(* IEC 61131-3 sources: ADRC_WWTP/PLC_ST/Codigos, 7 files *)

(* ---- ADRC_ESO.st ---- *)
FUNCTION_BLOCK ADRC_ESO
VAR_INPUT
    SET_POINT : LREAL;              (* setpoint r *)
    ACTUAL    : LREAL;              (* measurement y *)
    WC        : LREAL;              (* controller bandwidth [rad/s] *)
    WO        : LREAL;              (* observer bandwidth [rad/s] *)
    B0        : LREAL;              (* plant input gain *)
    TS        : TIME := T#50MS;     (* sampling time, equal to the task period *)
    U_MIN     : LREAL := 0.0;
    U_MAX     : LREAL := 100.0;
    RESET     : BOOL := FALSE;
END_VAR
VAR_OUTPUT
    U         : LREAL;              (* control signal to the actuator *)
END_VAR
VAR CONSTANT
    ST_RESET     : INT := 0;
    ST_AUTOMATIC : INT := 1;
END_VAR
VAR
    T_S       : LREAL;              (* sampling time [s] *)
    State     : INT;
    Ready     : BOOL := FALSE;      (* valid gains available *)
    A         : ARRAY[1..2, 1..2] OF LREAL;
    B         : ARRAY[1..2] OF LREAL;
    C         : ARRAY[1..2] OF LREAL;
    L         : ARRAY[1..2] OF LREAL;
    K         : ARRAY[1..2] OF LREAL;
    X         : ARRAY[1..2] OF LREAL;   (* x_hat: estimated error and total disturbance *)
    X_old     : ARRAY[1..2] OF LREAL;
    Ey, Ey_old : LREAL;
    U0, U0_old : LREAL;
    Bo, Zc, Zo : LREAL;
END_VAR

(* state selection *)
IF RESET OR NOT Ready THEN
    State := ST_RESET;
ELSE
    State := ST_AUTOMATIC;
END_IF

(* sampling time in seconds *)
T_S := TIME_TO_LREAL(TS) / 1000.0;

(* gains are only updated outside AUTOMATIC *)
IF (State <> ST_AUTOMATIC) AND (T_S > 0.0) AND (WC > 0.0) AND (WO > WC) AND (B0 > 0.0) THEN
    Zc := EXP(-WC * T_S);
    Zo := EXP(-WO * T_S);
    A[1,1] := 1.0;   A[1,2] := T_S;
    A[2,1] := 0.0;   A[2,2] := 1.0;
    B[1]   := T_S;    B[2]   := 0.0;
    C[1]   := 1.0;   C[2]   := 0.0;
    L[1]   := 2.0 * (1.0 - Zo);
    L[2]   := (1.0 - Zo) * (1.0 - Zo) / T_S;
    K[1]   := (1.0 - Zc) / T_S;
    K[2]   := 1.0;
    Bo     := B0;
    Ready  := TRUE;
END_IF

(* observer: x_hat[k] = (A - L C) x_hat[k-1] + B u0[k-1] + L ey[k-1] *)
X[1] := (A[1,1] - L[1]*C[1])*X_old[1] + (A[1,2] - L[1]*C[2])*X_old[2] + B[1]*U0_old + L[1]*Ey_old;
X[2] := (A[2,1] - L[2]*C[1])*X_old[1] + (A[2,2] - L[2]*C[2])*X_old[2] + B[2]*U0_old + L[2]*Ey_old;

CASE State OF
ST_RESET:
    (* output and observer to zero, as if it had just started *)
    U    := LIMIT(U_MIN, 0.0, U_MAX);
    X[1] := 0.0;
    X[2] := -Bo * U;
    Ey   := 0.0;

ST_AUTOMATIC:
    (* control law: u0 = -K x_hat[k],  u = u0/b0 *)
    Ey := ACTUAL - SET_POINT;
    U0 := -(K[1]*X[1] + K[2]*X[2]);
    U  := LIMIT(U_MIN, U0 / Bo, U_MAX);
END_CASE

(* the observer always receives the applied order *)
U0 := Bo * U;

X_old  := X;
U0_old := U0;
Ey_old := Ey;
END_FUNCTION_BLOCK

(* ---- ADRC_GPI.st ---- *)
FUNCTION_BLOCK ADRC_GPI
VAR_INPUT
    SET_POINT : LREAL;              (* setpoint r *)
    ACTUAL    : LREAL;              (* measurement y *)
    WC        : LREAL;              (* controller bandwidth [rad/s] *)
    WO        : LREAL;              (* observer bandwidth [rad/s] *)
    B0        : LREAL;              (* plant input gain *)
    TS        : TIME := T#50MS;     (* sampling time, equal to the task period *)
    U_MIN     : LREAL := 0.0;
    U_MAX     : LREAL := 100.0;
    RESET     : BOOL := FALSE;
END_VAR
VAR_OUTPUT
    U         : LREAL;              (* control signal to the actuator *)
END_VAR
VAR CONSTANT
    ST_RESET     : INT := 0;
    ST_AUTOMATIC : INT := 1;
END_VAR
VAR
    T_S       : LREAL;              (* sampling time [s] *)
    State     : INT;
    Ready     : BOOL := FALSE;      (* valid gains available *)
    Bo, D0, Q : LREAL;
    A1, A2    : LREAL;              (* common denominator of H1 and H2 *)
    B0z, B1z, B2z : LREAL;          (* numerator of H1 *)
    G0, G1, G2    : LREAL;          (* numerator of H2 *)
    E, E_1, E_2   : LREAL;          (* r - y and its delays *)
    V, V_1, V_2   : LREAL;
    U_1, U_2, W   : LREAL;
END_VAR

(* state selection *)
IF RESET OR NOT Ready THEN
    State := ST_RESET;
ELSE
    State := ST_AUTOMATIC;
END_IF

(* sampling time in seconds *)
T_S := TIME_TO_LREAL(TS) / 1000.0;

(* gains are only updated outside AUTOMATIC *)
IF (State <> ST_AUTOMATIC) AND (T_S > 0.0) AND (WC > 0.0) AND (WO > WC) AND (B0 > 0.0) THEN
    (* Tustin with E1(s) = (s + wo)^2 *)
    Q   := 2.0 + WO * T_S;
    D0  := Q * Q;
    A1  := -2.0 * (4.0 - WO * WO * T_S * T_S) / D0;
    A2  := (2.0 - WO * T_S) * (2.0 - WO * T_S) / D0;
    B0z := WO * T_S * (WC * WO * T_S + 2.0 * (WO + 2.0 * WC)) / D0;
    B1z := 2.0 * WC * WO * WO * T_S * T_S / D0;
    B2z := WO * T_S * (WC * WO * T_S - 2.0 * (WO + 2.0 * WC)) / D0;
    G0  := T_S * (2.0 * WC - WO * WO * T_S) / D0;
    G1  := -2.0 * WO * WO * T_S * T_S / D0;
    G2  := -T_S * (2.0 * WC + WO * WO * T_S) / D0;
    Bo  := B0;
    Ready := TRUE;
END_IF

CASE State OF
ST_RESET:
    (* output and delays to zero, as if it had just started *)
    U := LIMIT(U_MIN, 0.0, U_MAX);
    E := 0.0;   E_1 := 0.0;   E_2 := 0.0;
    V := U;     V_1 := U;     V_2 := U;
    U_1 := U;   U_2 := U;

ST_AUTOMATIC:
    (* direct form I; 1 + G0 solves the loop through the direct term of H2 *)
    E := SET_POINT - ACTUAL;
    W := (B0z*E + B1z*E_1 + B2z*E_2) / Bo - (G1*U_1 + G2*U_2) - A1*V_1 - A2*V_2;
    U := LIMIT(U_MIN, W / (1.0 + G0), U_MAX);
    V := W - G0 * U;
END_CASE

(* shift: oldest first *)
E_2 := E_1;   E_1 := E;
V_2 := V_1;   V_1 := V;
U_2 := U_1;   U_1 := U;
END_FUNCTION_BLOCK

(* ---- BEZIER_REF.st ---- *)
FUNCTION_BLOCK BEZIER_REF
VAR_INPUT
    SET_POINT : LREAL;              (* setpoint r *)
    ACTUAL    : LREAL;              (* measurement y *)
    TF        : TIME := T#20M;      (* segment duration, taken at each setpoint change *)
    TS        : TIME := T#50MS;     (* sampling time, equal to the task period *)
    RESET     : BOOL := FALSE;
END_VAR
VAR_OUTPUT
    Y         : LREAL;              (* reference y*, goes to the controller *)
END_VAR
VAR CONSTANT
    ST_RESET     : INT := 0;
    ST_AUTOMATIC : INT := 1;
END_VAR
VAR
    T_S       : LREAL;              (* sampling time [s] *)
    T_F       : LREAL;              (* segment duration [s] *)
    State     : INT;
    Ready     : BOOL := FALSE;      (* valid parameters available *)
    Ts_set         : LREAL;
    Tf_set         : LREAL;         (* duration of the current segment *)
    Yc, Dyc, Yf    : LREAL;         (* segment start state and target *)
    Delta, C1, C2, C3 : LREAL;      (* polynomial coefficients in tau *)
    Dy, Tn, Cnt, SP_old : LREAL;
END_VAR

(* state selection *)
IF RESET OR NOT Ready THEN
    State := ST_RESET;
ELSE
    State := ST_AUTOMATIC;
END_IF

(* times in seconds *)
T_S := TIME_TO_LREAL(TS) / 1000.0;
T_F := TIME_TO_LREAL(TF) / 1000.0;

(* parameters are only updated outside AUTOMATIC *)
IF (State <> ST_AUTOMATIC) AND (T_S > 0.0) AND (T_F > 0.0) THEN
    Ts_set := T_S;
    Tf_set := T_F;
    Ready  := TRUE;
END_IF

CASE State OF
ST_RESET:
    (* at rest on the measurement; leaving RESET starts the manoeuvre again *)
    Y  := ACTUAL;   Dy := 0.0;
    Yc := ACTUAL;   Dyc := 0.0;   Yf := ACTUAL;
    C1 := 0.0;      C2 := 0.0;    C3 := 0.0;
    Cnt := 0.0;     SP_old := ACTUAL;

ST_AUTOMATIC:
    (* evaluate the current segment, tau = n Ts/Tf *)
    Tn := Cnt * Ts_set / Tf_set;
    IF Tn < 1.0 THEN
        Y  := Yc + Tn * (C1 + Tn * (C2 + Tn * C3));
        Dy := (C1 + Tn * (2.0 * C2 + 3.0 * Tn * C3)) / Tf_set;
    ELSE
        Y  := Yf;
        Dy := 0.0;
    END_IF

    (* new setpoint: replan from the state of the reference *)
    IF SET_POINT <> SP_old THEN
        Yc := Y;
        Dyc := Dy;
        Yf := SET_POINT;
        Delta := Yf - Yc;
        IF T_F > 0.0 THEN
            Tf_set := T_F;
        END_IF
        C1 := Dyc * Tf_set;
        C2 := 3.0 * Delta - 2.0 * Dyc * Tf_set;
        C3 := -2.0 * Delta + Dyc * Tf_set;
        Cnt := 0.0;
        SP_old := SET_POINT;
    END_IF

    IF Cnt * Ts_set < Tf_set THEN
        Cnt := Cnt + 1.0;
    END_IF
END_CASE

END_FUNCTION_BLOCK

(* ---- GPI.st ---- *)
FUNCTION_BLOCK GPI
VAR_INPUT
    SET_POINT : LREAL;              (* setpoint r *)
    ACTUAL    : LREAL;              (* measurement y *)
    K0        : LREAL;              (* GPI gains: (k1 s + k0)/(s (s + k2)) *)
    K1        : LREAL;
    K2        : LREAL;
    B0        : LREAL;              (* plant input gain *)
    TS        : TIME := T#50MS;     (* sampling time, equal to the task period *)
    U_MIN     : LREAL := 0.0;
    U_MAX     : LREAL := 100.0;
    RESET     : BOOL := FALSE;
END_VAR
VAR_OUTPUT
    U         : LREAL;              (* control signal to the actuator *)
END_VAR
VAR CONSTANT
    ST_RESET     : INT := 0;
    ST_AUTOMATIC : INT := 1;
END_VAR
VAR
    T_S       : LREAL;              (* sampling time [s] *)
    State     : INT;
    Ready     : BOOL := FALSE;      (* valid gains available *)
    Bo, D0, Q : LREAL;
    A1, A2    : LREAL;              (* common denominator of H1 and H2 *)
    B0z, B1z, B2z : LREAL;          (* numerator of H1 *)
    G0, G1, G2    : LREAL;          (* numerator of H2 *)
    E, E_1, E_2   : LREAL;          (* r - y and its delays *)
    V, V_1, V_2   : LREAL;
    U_1, U_2, W   : LREAL;
END_VAR

(* state selection *)
IF RESET OR NOT Ready THEN
    State := ST_RESET;
ELSE
    State := ST_AUTOMATIC;
END_IF

(* sampling time in seconds *)
T_S := TIME_TO_LREAL(TS) / 1000.0;

(* gains are only updated outside AUTOMATIC, and only if they are stable *)
IF (State <> ST_AUTOMATIC) AND (T_S > 0.0) AND (B0 > 0.0) AND (K0 > 0.0) AND (K1 > 0.0)
        AND (K2 > 0.0) AND (K2 * K1 > K0) THEN
    (* Tustin with E1(s) = s^2 + k2 s + k1 *)
    Q   := K1 * T_S * T_S;
    D0  := 4.0 + 2.0 * K2 * T_S + Q;
    A1  := (2.0 * Q - 8.0) / D0;
    A2  := (4.0 - 2.0 * K2 * T_S + Q) / D0;
    B0z := (K0 * T_S * T_S + 2.0 * K1 * T_S) / D0;
    B1z := 2.0 * K0 * T_S * T_S / D0;
    B2z := (K0 * T_S * T_S - 2.0 * K1 * T_S) / D0;
    G0  := -Q / D0;
    G1  := -2.0 * Q / D0;
    G2  := -Q / D0;
    Bo  := B0;
    Ready := TRUE;
END_IF

CASE State OF
ST_RESET:
    (* output and delays to zero, as if it had just started *)
    U := LIMIT(U_MIN, 0.0, U_MAX);
    E := 0.0;   E_1 := 0.0;   E_2 := 0.0;
    V := U;     V_1 := U;     V_2 := U;
    U_1 := U;   U_2 := U;

ST_AUTOMATIC:
    (* direct form I; 1 + G0 solves the loop through the direct term of H2 *)
    E := SET_POINT - ACTUAL;
    W := (B0z*E + B1z*E_1 + B2z*E_2) / Bo - (G1*U_1 + G2*U_2) - A1*V_1 - A2*V_2;
    U := LIMIT(U_MIN, W / (1.0 + G0), U_MAX);
    V := W - G0 * U;
END_CASE

(* shift: oldest first *)
E_2 := E_1;   E_1 := E;
V_2 := V_1;   V_1 := V;
U_2 := U_1;   U_1 := U;
END_FUNCTION_BLOCK

(* ---- PLANT.st ---- *)
FUNCTION_BLOCK PLANT
VAR_INPUT
    U        : LREAL;               (* plant input *)
    K_DC     : LREAL;               (* DC gain *)
    TAU      : LREAL;               (* time constant [s] *)
    TS       : TIME := T#50MS;      (* sampling time, equal to the task period *)
END_VAR
VAR_OUTPUT
    Y        : LREAL;               (* plant output *)
END_VAR
VAR
    T_S      : LREAL;               (* sampling time [s] *)
    Ag, Bg   : LREAL;
    U_1      : LREAL;               (* previous input *)
END_VAR

(* sampling time in seconds *)
T_S := TIME_TO_LREAL(TS) / 1000.0;

(* first-order plant K_DC/(TAU s + 1), discretized with Tustin *)
Ag := (T_S - 2.0 * TAU) / (T_S + 2.0 * TAU);
Bg := K_DC * T_S / (T_S + 2.0 * TAU);

(* call it after the controller: Y is the next measurement *)
Y   := -Ag * Y + Bg * (U + U_1);
U_1 := U;
END_FUNCTION_BLOCK

(* ---- PREFILTER_ADRC.st ---- *)
FUNCTION_BLOCK PREFILTER_ADRC
VAR_INPUT
    SET_POINT : LREAL;              (* setpoint r *)
    ACTUAL    : LREAL;              (* measurement y *)
    WC        : LREAL;              (* controller bandwidth [rad/s] *)
    WO        : LREAL;              (* observer bandwidth [rad/s] *)
    TS        : TIME := T#50MS;     (* sampling time, equal to the task period *)
    RESET     : BOOL := FALSE;
END_VAR
VAR_OUTPUT
    Y         : LREAL;              (* filtered setpoint, goes to the controller *)
END_VAR
VAR CONSTANT
    ST_RESET     : INT := 0;
    ST_AUTOMATIC : INT := 1;
END_VAR
VAR
    T_S       : LREAL;              (* sampling time [s] *)
    State     : INT;
    Ready     : BOOL := FALSE;      (* valid gains available *)
    Af, Bf, Q : LREAL;
    Y_1, R_1  : LREAL;              (* delays of the output and the setpoint *)
END_VAR

(* state selection *)
IF RESET OR NOT Ready THEN
    State := ST_RESET;
ELSE
    State := ST_AUTOMATIC;
END_IF

(* sampling time in seconds *)
T_S := TIME_TO_LREAL(TS) / 1000.0;

(* gains are only updated outside AUTOMATIC *)
IF (State <> ST_AUTOMATIC) AND (T_S > 0.0) AND (WC > 0.0) AND (WO > WC) THEN
    (* Tustin of k0/(k1 s + k0), with k0/k1 = wc wo/(wo + 2 wc) *)
    Q  := 2.0 * (WO + 2.0 * WC);
    Af := (WC * WO * T_S - Q) / (WC * WO * T_S + Q);
    Bf := WC * WO * T_S / (WC * WO * T_S + Q);
    Ready := TRUE;
END_IF

CASE State OF
ST_RESET:
    (* follow the measurement; leaving RESET starts from it *)
    Y   := ACTUAL;
    Y_1 := ACTUAL;
    R_1 := ACTUAL;

ST_AUTOMATIC:
    (* r_f[k] = -af r_f[k-1] + bf (r[k] + r[k-1]) *)
    Y   := -Af * Y_1 + Bf * (SET_POINT + R_1);
    Y_1 := Y;
    R_1 := SET_POINT;
END_CASE

END_FUNCTION_BLOCK

(* ---- PREFILTER_GPI.st ---- *)
FUNCTION_BLOCK PREFILTER_GPI
VAR_INPUT
    SET_POINT : LREAL;              (* setpoint r *)
    ACTUAL    : LREAL;              (* measurement y *)
    K0        : LREAL;              (* prefilter: k0/(k1 s + k0) *)
    K1        : LREAL;
    TS        : TIME := T#50MS;     (* sampling time, equal to the task period *)
    RESET     : BOOL := FALSE;
END_VAR
VAR_OUTPUT
    Y         : LREAL;              (* filtered setpoint, goes to the controller *)
END_VAR
VAR CONSTANT
    ST_RESET     : INT := 0;
    ST_AUTOMATIC : INT := 1;
END_VAR
VAR
    T_S       : LREAL;              (* sampling time [s] *)
    State     : INT;
    Ready     : BOOL := FALSE;      (* valid gains available *)
    Af, Bf    : LREAL;
    Y_1, R_1  : LREAL;              (* delays of the output and the setpoint *)
END_VAR

(* state selection *)
IF RESET OR NOT Ready THEN
    State := ST_RESET;
ELSE
    State := ST_AUTOMATIC;
END_IF

(* sampling time in seconds *)
T_S := TIME_TO_LREAL(TS) / 1000.0;

(* gains are only updated outside AUTOMATIC *)
IF (State <> ST_AUTOMATIC) AND (T_S > 0.0) AND (K0 > 0.0) AND (K1 > 0.0) THEN
    (* Tustin *)
    Af := (K0 * T_S - 2.0 * K1) / (K0 * T_S + 2.0 * K1);
    Bf := K0 * T_S / (K0 * T_S + 2.0 * K1);
    Ready := TRUE;
END_IF

CASE State OF
ST_RESET:
    (* follow the measurement; leaving RESET starts from it *)
    Y   := ACTUAL;
    Y_1 := ACTUAL;
    R_1 := ACTUAL;

ST_AUTOMATIC:
    (* r_f[k] = -af r_f[k-1] + bf (r[k] + r[k-1]) *)
    Y   := -Af * Y_1 + Bf * (SET_POINT + R_1);
    Y_1 := Y;
    R_1 := SET_POINT;
END_CASE

END_FUNCTION_BLOCK
